Fanuc KAREL source: KD00008.KL

PROGRAM KD00008
%NOLOCKGROUP
%TPMOTION
VAR
  I: INTEGER
  J: INTEGER
  B: BOOLEAN
  R: REAL
  S: STRING[80]
BEGIN
  I = 1
END KD00008
